Fanuc KAREL source: KT00385.KL

PROGRAM KT00385
%NOLOCKGROUP
VAR
  P1: POSITION
  P2: XYZWPREXT
  OUT: BOOLEAN
BEGIN
    P2.Y = 2.0
  OUT = P1 <= P2
END KT00385
